VAR_GLOBAL
		(*----------------> Real Time Clock <------------------*)

	dtRealTime								:DATE_AND_TIME;
	sRealTime								:STRING[22];
	stSystemTime							:TimeStruct;
	stSystemTime_Empty						:TimeStruct;
	sDateShort								:STRING[20];	(*	YYMMDD	*)
	
(*..........................................................................System TIME.....................................................................................*)
	sTime					: STRING[20];
	sDate					: STRING[20];
	sDateTime				: STRING[60];
	sTimeWithMicroSec		: STRING[40];

END_VAR

(* stored: Version 1.1.0.1, ProductVersion 3.1.4024.15
   GVL GVL_Time_12: Id {d439de53-09ae-4ded-89f7-367941b19f70} *)
